Fanuc KAREL source: KB00078.KL

PROGRAM KB00078
%NOLOCKGROUP
%ENVIRONMENT FLBT
VAR
  P1: FILE
  RESULT: INTEGER
BEGIN
  RESULT = GET_FILE_POS(P1)
END KB00078
